(* IEC 61131-3 sources: SRCI_CLIENT_PLC/RobotLibrary/Library/Structures/Telegram/PlcToRob/Command, 2 files *)

(* ---- TelegramPlcToRobCommand.st ---- *)
{attribute 'pack_mode' := '1'}
// -------------------------------------------------------------------------
//  SRCI Robot Library
// -------------------------------------------------------------------------
//
//  Object:      TelegramPlcToRobMessage
//  Author:      Thorsten Brach
//  Date:        2024-06-01
//
//  Description:
//
//
//  Copyright:
//    (C) 2024 Thorsten Brach. All rights reserved
//             Licensed under the MIT License.
//
//  Disclaimer:
//    This project is provided without any guarantee and can be used for
//    private and commercial purposes. Any use is at the user’s
//    own risk and responsibility.
//
// -------------------------------------------------------------------------
TYPE TelegramPlcToRobCommand :
STRUCT
  /// Header
  Header  : TelegramPlcToRobCommandHeader;
  /// Payload
  Payload : ARRAY[0..RobotLibraryParameter.PARAMETER_PAYLOAD_MAX] OF BYTE;
END_STRUCT
END_TYPE

(* ---- TelegramPlcToRobCommandHeader.st ---- *)
{attribute 'pack_mode' := '1'}
// -------------------------------------------------------------------------
//  SRCI Robot Library
// -------------------------------------------------------------------------
//
//  Object:      TelegramPlcToRobMessageHeader
//  Author:      Thorsten Brach
//  Date:        2024-06-01
//
//  Description:
//
//
//  Copyright:
//    (C) 2024 Thorsten Brach. All rights reserved
//             Licensed under the MIT License.
//
//  Disclaimer:
//    This project is provided without any guarantee and can be used for
//    private and commercial purposes. Any use is at the user’s
//    own risk and responsibility.
//
// -------------------------------------------------------------------------
TYPE TelegramPlcToRobCommandHeader :
STRUCT
  /// Command type
  CmdType           : CmdType;
  /// CMD priority level
  Prio              : PriorityLevel;
  /// Execution Mode
  ExecMode          : ExecutionMode;
  /// Parameter Sequence
  ParSequence       : BYTE;
END_STRUCT
END_TYPE
